(* IEC 61131-3 sources: stateaware-ics-monitoring/tests/st_gen/golden/ctown, 9 files *)

(* ---- ctown_plc1.st ---- *)
(* Auto-generated by st_gen 0.1.0 from ctown.inp + ctown_plcs.yaml
   Topology: ctown   PLC: PLC1
   SURROGATE Structured Text: reconstructed by st_gen from the EPANET INP model
   and a DHALSIM-style plcs.yaml. This is NOT the original vendor or benchmark
   PLC source code and must not be presented as such.
   Upstream: DHALSIM https://github.com/Critical-Infrastructure-Systems-Lab/DHALSIM @ 51a5e00f65cdd666b9aec10d3c928ea40ad1b53d
   DO NOT EDIT. *)

PROGRAM PLC1
VAR_INPUT
    T1 : REAL;            (* sourced from PLC2 *)
END_VAR
VAR_OUTPUT
    PU1 : BOOL;
    PU2 : BOOL;
END_VAR
VAR
    PU1_State : INT := 0;
    PU2_State : INT := 1;
END_VAR

(* ----- FSM for actuator PU1 ----- *)
CASE PU1_State OF
    0:  (* CLOSED *)
        PU1 := FALSE;
        IF T1 < 4 THEN
            PU1_State := 1;
        END_IF;
    1:  (* OPEN *)
        PU1 := TRUE;
        IF T1 > 6.3 THEN
            PU1_State := 0;
        END_IF;
END_CASE;

(* ----- FSM for actuator PU2 ----- *)
CASE PU2_State OF
    0:  (* CLOSED *)
        PU2 := FALSE;
        IF T1 < 1 THEN
            PU2_State := 1;
        END_IF;
    1:  (* OPEN *)
        PU2 := TRUE;
        IF T1 > 4.5 THEN
            PU2_State := 0;
        END_IF;
END_CASE;

END_PROGRAM

(* ---- ctown_plc2.st ---- *)
(* Auto-generated by st_gen 0.1.0 from ctown.inp + ctown_plcs.yaml
   Topology: ctown   PLC: PLC2
   SURROGATE Structured Text: reconstructed by st_gen from the EPANET INP model
   and a DHALSIM-style plcs.yaml. This is NOT the original vendor or benchmark
   PLC source code and must not be presented as such.
   Upstream: DHALSIM https://github.com/Critical-Infrastructure-Systems-Lab/DHALSIM @ 51a5e00f65cdd666b9aec10d3c928ea40ad1b53d
   DO NOT EDIT. *)

PROGRAM PLC2
(* No actuators with [CONTROLS] entries -- sensor-only or static-setting PLC. *)
END_PROGRAM

(* ---- ctown_plc3.st ---- *)
(* Auto-generated by st_gen 0.1.0 from ctown.inp + ctown_plcs.yaml
   Topology: ctown   PLC: PLC3
   SURROGATE Structured Text: reconstructed by st_gen from the EPANET INP model
   and a DHALSIM-style plcs.yaml. This is NOT the original vendor or benchmark
   PLC source code and must not be presented as such.
   Upstream: DHALSIM https://github.com/Critical-Infrastructure-Systems-Lab/DHALSIM @ 51a5e00f65cdd666b9aec10d3c928ea40ad1b53d
   DO NOT EDIT. *)

PROGRAM PLC3
VAR_INPUT
    T2 : REAL;            (* owned by this PLC *)
    T3 : REAL;            (* sourced from PLC4 *)
    T4 : REAL;            (* sourced from PLC6 *)
END_VAR
VAR_OUTPUT
    V2 : BOOL;
    PU4 : BOOL;
    PU5 : BOOL;
    PU6 : BOOL;
    PU7 : BOOL;
END_VAR
VAR
    V2_State : INT := 0;
    PU4_State : INT := 0;
    PU5_State : INT := 0;
    PU6_State : INT := 0;
    PU7_State : INT := 0;
END_VAR

(* ----- FSM for actuator V2 ----- *)
CASE V2_State OF
    0:  (* CLOSED *)
        V2 := FALSE;
        IF T2 < 0.5 THEN
            V2_State := 1;
        END_IF;
    1:  (* OPEN *)
        V2 := TRUE;
        IF T2 > 5.5 THEN
            V2_State := 0;
        END_IF;
END_CASE;

(* ----- FSM for actuator PU4 ----- *)
CASE PU4_State OF
    0:  (* CLOSED *)
        PU4 := FALSE;
        IF T3 < 3 THEN
            PU4_State := 1;
        END_IF;
    1:  (* OPEN *)
        PU4 := TRUE;
        IF T3 > 5.3 THEN
            PU4_State := 0;
        END_IF;
END_CASE;

(* ----- FSM for actuator PU5 ----- *)
CASE PU5_State OF
    0:  (* CLOSED *)
        PU5 := FALSE;
        IF T3 < 1 THEN
            PU5_State := 1;
        END_IF;
    1:  (* OPEN *)
        PU5 := TRUE;
        IF T3 > 3.5 THEN
            PU5_State := 0;
        END_IF;
END_CASE;

(* ----- FSM for actuator PU6 ----- *)
CASE PU6_State OF
    0:  (* CLOSED *)
        PU6 := FALSE;
        IF T4 < 2 THEN
            PU6_State := 1;
        END_IF;
    1:  (* OPEN *)
        PU6 := TRUE;
        IF T4 > 3.5 THEN
            PU6_State := 0;
        END_IF;
END_CASE;

(* ----- FSM for actuator PU7 ----- *)
CASE PU7_State OF
    0:  (* CLOSED *)
        PU7 := FALSE;
        IF T4 < 3 THEN
            PU7_State := 1;
        END_IF;
    1:  (* OPEN *)
        PU7 := TRUE;
        IF T4 > 4.5 THEN
            PU7_State := 0;
        END_IF;
END_CASE;

END_PROGRAM

(* ---- ctown_plc4.st ---- *)
(* Auto-generated by st_gen 0.1.0 from ctown.inp + ctown_plcs.yaml
   Topology: ctown   PLC: PLC4
   SURROGATE Structured Text: reconstructed by st_gen from the EPANET INP model
   and a DHALSIM-style plcs.yaml. This is NOT the original vendor or benchmark
   PLC source code and must not be presented as such.
   Upstream: DHALSIM https://github.com/Critical-Infrastructure-Systems-Lab/DHALSIM @ 51a5e00f65cdd666b9aec10d3c928ea40ad1b53d
   DO NOT EDIT. *)

PROGRAM PLC4
(* No actuators with [CONTROLS] entries -- sensor-only or static-setting PLC. *)
END_PROGRAM

(* ---- ctown_plc5.st ---- *)
(* Auto-generated by st_gen 0.1.0 from ctown.inp + ctown_plcs.yaml
   Topology: ctown   PLC: PLC5
   SURROGATE Structured Text: reconstructed by st_gen from the EPANET INP model
   and a DHALSIM-style plcs.yaml. This is NOT the original vendor or benchmark
   PLC source code and must not be presented as such.
   Upstream: DHALSIM https://github.com/Critical-Infrastructure-Systems-Lab/DHALSIM @ 51a5e00f65cdd666b9aec10d3c928ea40ad1b53d
   DO NOT EDIT. *)

PROGRAM PLC5
VAR_INPUT
    T5 : REAL;            (* sourced from PLC7 *)
    T7 : REAL;            (* sourced from PLC9 *)
END_VAR
VAR_OUTPUT
    PU8 : BOOL;
    PU10 : BOOL;
    PU11 : BOOL;
END_VAR
VAR
    PU8_State : INT := 0;
    PU10_State : INT := 0;
    PU11_State : INT := 0;
END_VAR

(* ----- FSM for actuator PU8 ----- *)
CASE PU8_State OF
    0:  (* CLOSED *)
        PU8 := FALSE;
        IF T5 < 1.5 THEN
            PU8_State := 1;
        END_IF;
    1:  (* OPEN *)
        PU8 := TRUE;
        IF T5 > 4 THEN
            PU8_State := 0;
        END_IF;
END_CASE;

(* ----- FSM for actuator PU10 ----- *)
CASE PU10_State OF
    0:  (* CLOSED *)
        PU10 := FALSE;
        IF T7 < 1.5 THEN
            PU10_State := 1;
        END_IF;
    1:  (* OPEN *)
        PU10 := TRUE;
        IF T7 > 4.8 THEN
            PU10_State := 0;
        END_IF;
END_CASE;

(* ----- FSM for actuator PU11 ----- *)
CASE PU11_State OF
    0:  (* CLOSED *)
        PU11 := FALSE;
        IF T7 < 0.5 THEN
            PU11_State := 1;
        END_IF;
    1:  (* OPEN *)
        PU11 := TRUE;
        IF T7 > 3 THEN
            PU11_State := 0;
        END_IF;
END_CASE;

END_PROGRAM

(* ---- ctown_plc6.st ---- *)
(* Auto-generated by st_gen 0.1.0 from ctown.inp + ctown_plcs.yaml
   Topology: ctown   PLC: PLC6
   SURROGATE Structured Text: reconstructed by st_gen from the EPANET INP model
   and a DHALSIM-style plcs.yaml. This is NOT the original vendor or benchmark
   PLC source code and must not be presented as such.
   Upstream: DHALSIM https://github.com/Critical-Infrastructure-Systems-Lab/DHALSIM @ 51a5e00f65cdd666b9aec10d3c928ea40ad1b53d
   DO NOT EDIT. *)

PROGRAM PLC6
(* No actuators with [CONTROLS] entries -- sensor-only or static-setting PLC. *)
END_PROGRAM

(* ---- ctown_plc7.st ---- *)
(* Auto-generated by st_gen 0.1.0 from ctown.inp + ctown_plcs.yaml
   Topology: ctown   PLC: PLC7
   SURROGATE Structured Text: reconstructed by st_gen from the EPANET INP model
   and a DHALSIM-style plcs.yaml. This is NOT the original vendor or benchmark
   PLC source code and must not be presented as such.
   Upstream: DHALSIM https://github.com/Critical-Infrastructure-Systems-Lab/DHALSIM @ 51a5e00f65cdd666b9aec10d3c928ea40ad1b53d
   DO NOT EDIT. *)

PROGRAM PLC7
(* No actuators with [CONTROLS] entries -- sensor-only or static-setting PLC. *)
END_PROGRAM

(* ---- ctown_plc8.st ---- *)
(* Auto-generated by st_gen 0.1.0 from ctown.inp + ctown_plcs.yaml
   Topology: ctown   PLC: PLC8
   SURROGATE Structured Text: reconstructed by st_gen from the EPANET INP model
   and a DHALSIM-style plcs.yaml. This is NOT the original vendor or benchmark
   PLC source code and must not be presented as such.
   Upstream: DHALSIM https://github.com/Critical-Infrastructure-Systems-Lab/DHALSIM @ 51a5e00f65cdd666b9aec10d3c928ea40ad1b53d
   DO NOT EDIT. *)

PROGRAM PLC8
(* No actuators with [CONTROLS] entries -- sensor-only or static-setting PLC. *)
END_PROGRAM

(* ---- ctown_plc9.st ---- *)
(* Auto-generated by st_gen 0.1.0 from ctown.inp + ctown_plcs.yaml
   Topology: ctown   PLC: PLC9
   SURROGATE Structured Text: reconstructed by st_gen from the EPANET INP model
   and a DHALSIM-style plcs.yaml. This is NOT the original vendor or benchmark
   PLC source code and must not be presented as such.
   Upstream: DHALSIM https://github.com/Critical-Infrastructure-Systems-Lab/DHALSIM @ 51a5e00f65cdd666b9aec10d3c928ea40ad1b53d
   DO NOT EDIT. *)

PROGRAM PLC9
(* No actuators with [CONTROLS] entries -- sensor-only or static-setting PLC. *)
END_PROGRAM
